// TIA Portal V19 export
FUNCTION "MB_VFD" : Void   // FC1, LAD
{ S7_Optimized_Access := 'TRUE' }
// stored: SetENOAutomatically false
   VAR_TEMP   // added for the SCL form of the ladder/FBD networks
      _w1 : Bool;
   END_VAR
BEGIN

REGION Network 1
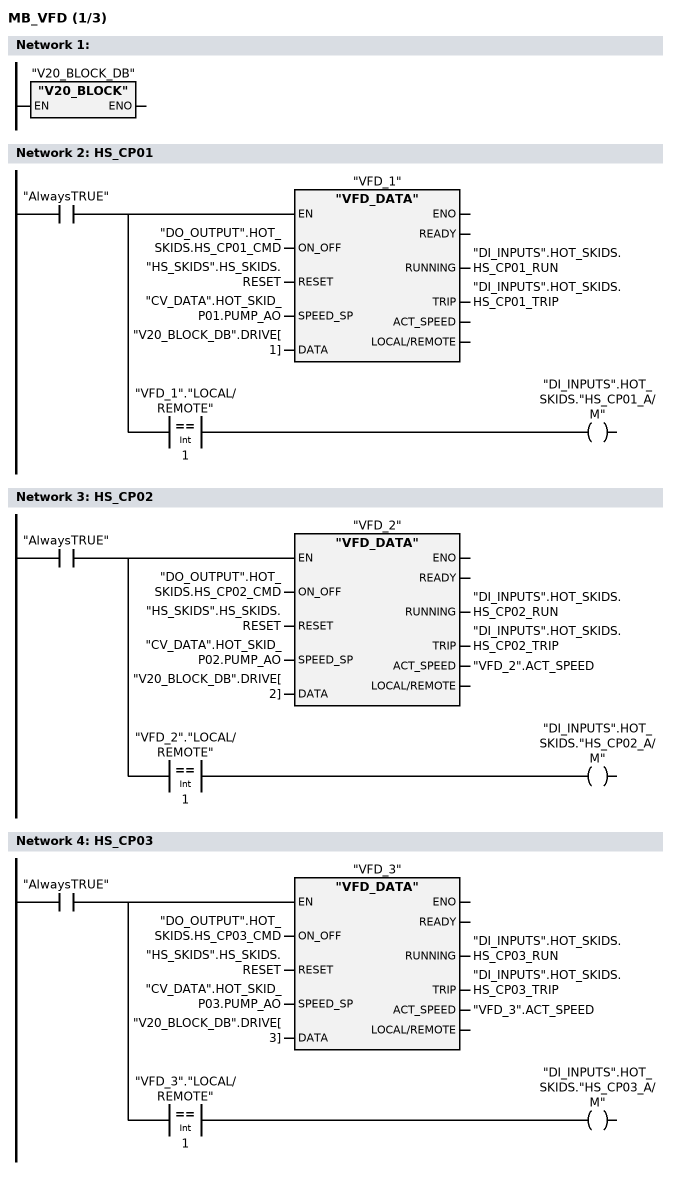
   RUNG wire#powerrail
      "V20_BLOCK_DB"()
   END_RUNG
   // the same network as SCL:
   "V20_BLOCK_DB"();   // "V20_BLOCK"
END_REGION

REGION Network 2: HS_CP01
   RUNG wire#powerrail
      Contact( "AlwaysTRUE" )
      wire#w1
      "VFD_1"(ON_OFF := "DO_OUTPUT".HOT_SKIDS.HS_CP01_CMD, RESET := "HS_SKIDS".HS_SKIDS.RESET, SPEED_SP := "CV_DATA".HOT_SKID_P01.PUMP_AO, DATA := "V20_BLOCK_DB".DRIVE[1], READY =>, RUNNING => "DI_INPUTS".HOT_SKIDS.HS_CP01_RUN, TRIP => "DI_INPUTS".HOT_SKIDS.HS_CP01_TRIP, ACT_SPEED =>, "LOCAL/REMOTE" =>)
   END_RUNG
   RUNG wire#w1
      { S7_Templates := "SrcType := Int" } EQ_Contact(in1 := "VFD_1"."LOCAL/REMOTE", in2 := 1)
      Coil( "DI_INPUTS".HOT_SKIDS."HS_CP01_A/M" )
   END_RUNG
   // the same network as SCL:
   #_w1 := "AlwaysTRUE";
   IF #_w1 THEN
       "VFD_1"(ON_OFF := "DO_OUTPUT".HOT_SKIDS.HS_CP01_CMD,   // "VFD_DATA"
               RESET := "HS_SKIDS".HS_SKIDS.RESET,
               SPEED_SP := "CV_DATA".HOT_SKID_P01.PUMP_AO,
               DATA := "V20_BLOCK_DB".DRIVE[1],
               RUNNING => "DI_INPUTS".HOT_SKIDS.HS_CP01_RUN,
               TRIP => "DI_INPUTS".HOT_SKIDS.HS_CP01_TRIP);
   END_IF;
   "DI_INPUTS".HOT_SKIDS."HS_CP01_A/M" := #_w1 AND ("VFD_1"."LOCAL/REMOTE" = 1);
END_REGION

REGION Network 3: HS_CP02
   RUNG wire#powerrail
      Contact( "AlwaysTRUE" )
      wire#w1
      "VFD_2"(ON_OFF := "DO_OUTPUT".HOT_SKIDS.HS_CP02_CMD, RESET := "HS_SKIDS".HS_SKIDS.RESET, SPEED_SP := "CV_DATA".HOT_SKID_P02.PUMP_AO, DATA := "V20_BLOCK_DB".DRIVE[2], READY =>, RUNNING => "DI_INPUTS".HOT_SKIDS.HS_CP02_RUN, TRIP => "DI_INPUTS".HOT_SKIDS.HS_CP02_TRIP, ACT_SPEED => "VFD_2".ACT_SPEED, "LOCAL/REMOTE" =>)
   END_RUNG
   RUNG wire#w1
      { S7_Templates := "SrcType := Int" } EQ_Contact(in1 := "VFD_2"."LOCAL/REMOTE", in2 := 1)
      Coil( "DI_INPUTS".HOT_SKIDS."HS_CP02_A/M" )
   END_RUNG
   // the same network as SCL:
   #_w1 := "AlwaysTRUE";
   IF #_w1 THEN
       "VFD_2"(ON_OFF := "DO_OUTPUT".HOT_SKIDS.HS_CP02_CMD,   // "VFD_DATA"
               RESET := "HS_SKIDS".HS_SKIDS.RESET,
               SPEED_SP := "CV_DATA".HOT_SKID_P02.PUMP_AO,
               DATA := "V20_BLOCK_DB".DRIVE[2],
               RUNNING => "DI_INPUTS".HOT_SKIDS.HS_CP02_RUN,
               TRIP => "DI_INPUTS".HOT_SKIDS.HS_CP02_TRIP,
               ACT_SPEED => "VFD_2".ACT_SPEED);
   END_IF;
   "DI_INPUTS".HOT_SKIDS."HS_CP02_A/M" := #_w1 AND ("VFD_2"."LOCAL/REMOTE" = 1);
END_REGION

REGION Network 4: HS_CP03
   RUNG wire#powerrail
      Contact( "AlwaysTRUE" )
      wire#w1
      "VFD_3"(ON_OFF := "DO_OUTPUT".HOT_SKIDS.HS_CP03_CMD, RESET := "HS_SKIDS".HS_SKIDS.RESET, SPEED_SP := "CV_DATA".HOT_SKID_P03.PUMP_AO, DATA := "V20_BLOCK_DB".DRIVE[3], READY =>, RUNNING => "DI_INPUTS".HOT_SKIDS.HS_CP03_RUN, TRIP => "DI_INPUTS".HOT_SKIDS.HS_CP03_TRIP, ACT_SPEED => "VFD_3".ACT_SPEED, "LOCAL/REMOTE" =>)
   END_RUNG
   RUNG wire#w1
      { S7_Templates := "SrcType := Int" } EQ_Contact(in1 := "VFD_3"."LOCAL/REMOTE", in2 := 1)
      Coil( "DI_INPUTS".HOT_SKIDS."HS_CP03_A/M" )
   END_RUNG
   // the same network as SCL:
   #_w1 := "AlwaysTRUE";
   IF #_w1 THEN
       "VFD_3"(ON_OFF := "DO_OUTPUT".HOT_SKIDS.HS_CP03_CMD,   // "VFD_DATA"
               RESET := "HS_SKIDS".HS_SKIDS.RESET,
               SPEED_SP := "CV_DATA".HOT_SKID_P03.PUMP_AO,
               DATA := "V20_BLOCK_DB".DRIVE[3],
               RUNNING => "DI_INPUTS".HOT_SKIDS.HS_CP03_RUN,
               TRIP => "DI_INPUTS".HOT_SKIDS.HS_CP03_TRIP,
               ACT_SPEED => "VFD_3".ACT_SPEED);
   END_IF;
   "DI_INPUTS".HOT_SKIDS."HS_CP03_A/M" := #_w1 AND ("VFD_3"."LOCAL/REMOTE" = 1);
END_REGION

REGION Network 5: CHS_CP01
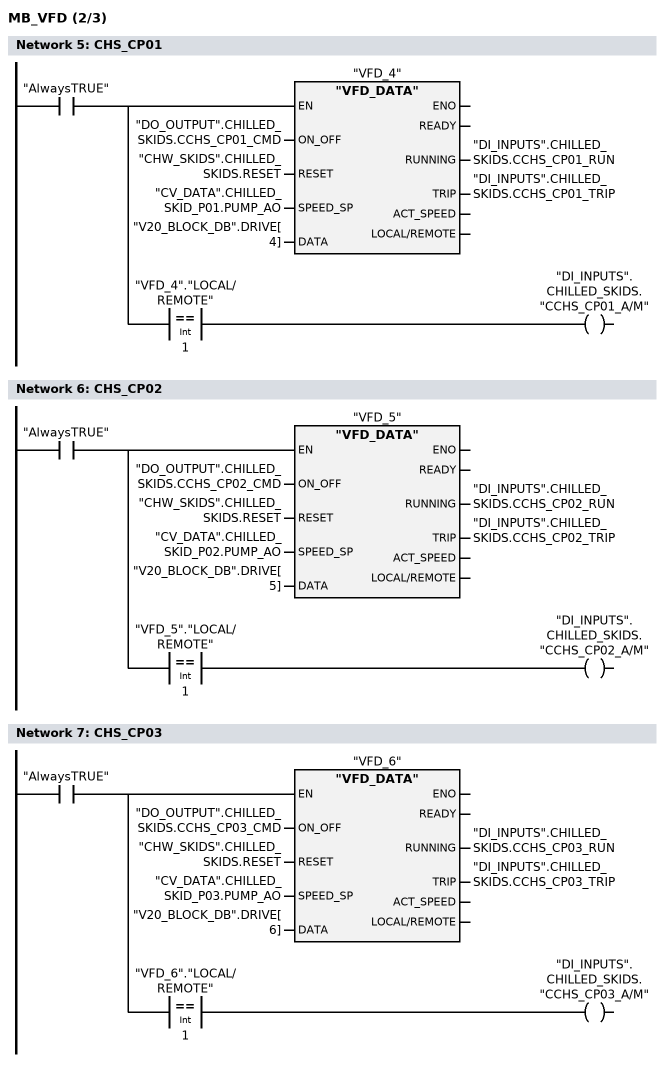
   RUNG wire#powerrail
      Contact( "AlwaysTRUE" )
      wire#w1
      "VFD_4"(ON_OFF := "DO_OUTPUT".CHILLED_SKIDS.CCHS_CP01_CMD, RESET := "CHW_SKIDS".CHILLED_SKIDS.RESET, SPEED_SP := "CV_DATA".CHILLED_SKID_P01.PUMP_AO, DATA := "V20_BLOCK_DB".DRIVE[4], READY =>, RUNNING => "DI_INPUTS".CHILLED_SKIDS.CCHS_CP01_RUN, TRIP => "DI_INPUTS".CHILLED_SKIDS.CCHS_CP01_TRIP, ACT_SPEED =>, "LOCAL/REMOTE" =>)
   END_RUNG
   RUNG wire#w1
      { S7_Templates := "SrcType := Int" } EQ_Contact(in1 := "VFD_4"."LOCAL/REMOTE", in2 := 1)
      Coil( "DI_INPUTS".CHILLED_SKIDS."CCHS_CP01_A/M" )
   END_RUNG
   // the same network as SCL:
   #_w1 := "AlwaysTRUE";
   IF #_w1 THEN
       "VFD_4"(ON_OFF := "DO_OUTPUT".CHILLED_SKIDS.CCHS_CP01_CMD,   // "VFD_DATA"
               RESET := "CHW_SKIDS".CHILLED_SKIDS.RESET,
               SPEED_SP := "CV_DATA".CHILLED_SKID_P01.PUMP_AO,
               DATA := "V20_BLOCK_DB".DRIVE[4],
               RUNNING => "DI_INPUTS".CHILLED_SKIDS.CCHS_CP01_RUN,
               TRIP => "DI_INPUTS".CHILLED_SKIDS.CCHS_CP01_TRIP);
   END_IF;
   "DI_INPUTS".CHILLED_SKIDS."CCHS_CP01_A/M" := #_w1 AND ("VFD_4"."LOCAL/REMOTE" = 1);
END_REGION

REGION Network 6: CHS_CP02
   RUNG wire#powerrail
      Contact( "AlwaysTRUE" )
      wire#w1
      "VFD_5"(ON_OFF := "DO_OUTPUT".CHILLED_SKIDS.CCHS_CP02_CMD, RESET := "CHW_SKIDS".CHILLED_SKIDS.RESET, SPEED_SP := "CV_DATA".CHILLED_SKID_P02.PUMP_AO, DATA := "V20_BLOCK_DB".DRIVE[5], READY =>, RUNNING => "DI_INPUTS".CHILLED_SKIDS.CCHS_CP02_RUN, TRIP => "DI_INPUTS".CHILLED_SKIDS.CCHS_CP02_TRIP, ACT_SPEED =>, "LOCAL/REMOTE" =>)
   END_RUNG
   RUNG wire#w1
      { S7_Templates := "SrcType := Int" } EQ_Contact(in1 := "VFD_5"."LOCAL/REMOTE", in2 := 1)
      Coil( "DI_INPUTS".CHILLED_SKIDS."CCHS_CP02_A/M" )
   END_RUNG
   // the same network as SCL:
   #_w1 := "AlwaysTRUE";
   IF #_w1 THEN
       "VFD_5"(ON_OFF := "DO_OUTPUT".CHILLED_SKIDS.CCHS_CP02_CMD,   // "VFD_DATA"
               RESET := "CHW_SKIDS".CHILLED_SKIDS.RESET,
               SPEED_SP := "CV_DATA".CHILLED_SKID_P02.PUMP_AO,
               DATA := "V20_BLOCK_DB".DRIVE[5],
               RUNNING => "DI_INPUTS".CHILLED_SKIDS.CCHS_CP02_RUN,
               TRIP => "DI_INPUTS".CHILLED_SKIDS.CCHS_CP02_TRIP);
   END_IF;
   "DI_INPUTS".CHILLED_SKIDS."CCHS_CP02_A/M" := #_w1 AND ("VFD_5"."LOCAL/REMOTE" = 1);
END_REGION

REGION Network 7: CHS_CP03
   RUNG wire#powerrail
      Contact( "AlwaysTRUE" )
      wire#w1
      "VFD_6"(ON_OFF := "DO_OUTPUT".CHILLED_SKIDS.CCHS_CP03_CMD, RESET := "CHW_SKIDS".CHILLED_SKIDS.RESET, SPEED_SP := "CV_DATA".CHILLED_SKID_P03.PUMP_AO, DATA := "V20_BLOCK_DB".DRIVE[6], READY =>, RUNNING => "DI_INPUTS".CHILLED_SKIDS.CCHS_CP03_RUN, TRIP => "DI_INPUTS".CHILLED_SKIDS.CCHS_CP03_TRIP, ACT_SPEED =>, "LOCAL/REMOTE" =>)
   END_RUNG
   RUNG wire#w1
      { S7_Templates := "SrcType := Int" } EQ_Contact(in1 := "VFD_6"."LOCAL/REMOTE", in2 := 1)
      Coil( "DI_INPUTS".CHILLED_SKIDS."CCHS_CP03_A/M" )
   END_RUNG
   // the same network as SCL:
   #_w1 := "AlwaysTRUE";
   IF #_w1 THEN
       "VFD_6"(ON_OFF := "DO_OUTPUT".CHILLED_SKIDS.CCHS_CP03_CMD,   // "VFD_DATA"
               RESET := "CHW_SKIDS".CHILLED_SKIDS.RESET,
               SPEED_SP := "CV_DATA".CHILLED_SKID_P03.PUMP_AO,
               DATA := "V20_BLOCK_DB".DRIVE[6],
               RUNNING => "DI_INPUTS".CHILLED_SKIDS.CCHS_CP03_RUN,
               TRIP => "DI_INPUTS".CHILLED_SKIDS.CCHS_CP03_TRIP);
   END_IF;
   "DI_INPUTS".CHILLED_SKIDS."CCHS_CP03_A/M" := #_w1 AND ("VFD_6"."LOCAL/REMOTE" = 1);
END_REGION

REGION Network 8: UCHS_CP01
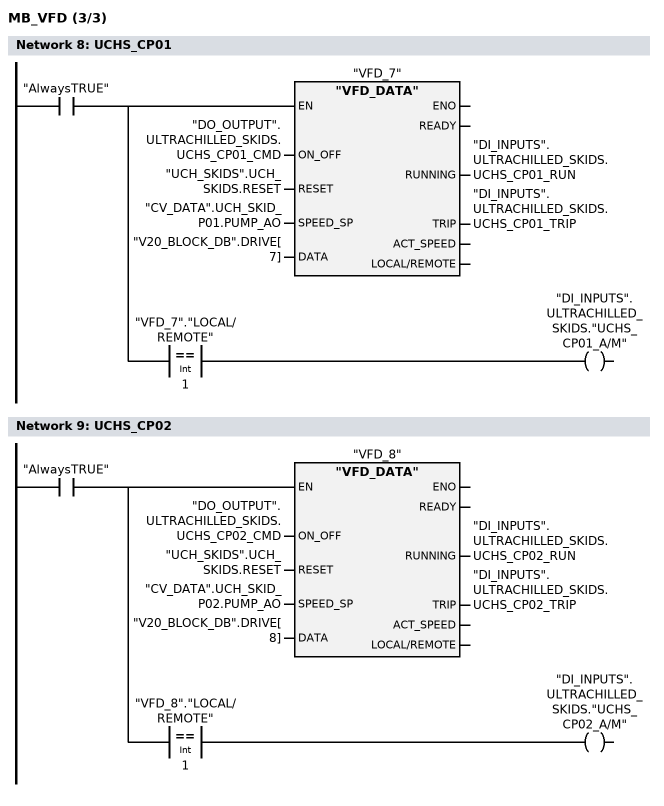
   RUNG wire#powerrail
      Contact( "AlwaysTRUE" )
      wire#w1
      "VFD_7"(ON_OFF := "DO_OUTPUT".ULTRACHILLED_SKIDS.UCHS_CP01_CMD, RESET := "UCH_SKIDS".UCH_SKIDS.RESET, SPEED_SP := "CV_DATA".UCH_SKID_P01.PUMP_AO, DATA := "V20_BLOCK_DB".DRIVE[7], READY =>, RUNNING => "DI_INPUTS".ULTRACHILLED_SKIDS.UCHS_CP01_RUN, TRIP => "DI_INPUTS".ULTRACHILLED_SKIDS.UCHS_CP01_TRIP, ACT_SPEED =>, "LOCAL/REMOTE" =>)
   END_RUNG
   RUNG wire#w1
      { S7_Templates := "SrcType := Int" } EQ_Contact(in1 := "VFD_7"."LOCAL/REMOTE", in2 := 1)
      Coil( "DI_INPUTS".ULTRACHILLED_SKIDS."UCHS_CP01_A/M" )
   END_RUNG
   // the same network as SCL:
   #_w1 := "AlwaysTRUE";
   IF #_w1 THEN
       "VFD_7"(ON_OFF := "DO_OUTPUT".ULTRACHILLED_SKIDS.UCHS_CP01_CMD,   // "VFD_DATA"
               RESET := "UCH_SKIDS".UCH_SKIDS.RESET,
               SPEED_SP := "CV_DATA".UCH_SKID_P01.PUMP_AO,
               DATA := "V20_BLOCK_DB".DRIVE[7],
               RUNNING => "DI_INPUTS".ULTRACHILLED_SKIDS.UCHS_CP01_RUN,
               TRIP => "DI_INPUTS".ULTRACHILLED_SKIDS.UCHS_CP01_TRIP);
   END_IF;
   "DI_INPUTS".ULTRACHILLED_SKIDS."UCHS_CP01_A/M" := #_w1 AND ("VFD_7"."LOCAL/REMOTE" = 1);
END_REGION

REGION Network 9: UCHS_CP02
   RUNG wire#powerrail
      Contact( "AlwaysTRUE" )
      wire#w1
      "VFD_8"(ON_OFF := "DO_OUTPUT".ULTRACHILLED_SKIDS.UCHS_CP02_CMD, RESET := "UCH_SKIDS".UCH_SKIDS.RESET, SPEED_SP := "CV_DATA".UCH_SKID_P02.PUMP_AO, DATA := "V20_BLOCK_DB".DRIVE[8], READY =>, RUNNING => "DI_INPUTS".ULTRACHILLED_SKIDS.UCHS_CP02_RUN, TRIP => "DI_INPUTS".ULTRACHILLED_SKIDS.UCHS_CP02_TRIP, ACT_SPEED =>, "LOCAL/REMOTE" =>)
   END_RUNG
   RUNG wire#w1
      { S7_Templates := "SrcType := Int" } EQ_Contact(in1 := "VFD_8"."LOCAL/REMOTE", in2 := 1)
      Coil( "DI_INPUTS".ULTRACHILLED_SKIDS."UCHS_CP02_A/M" )
   END_RUNG
   // the same network as SCL:
   #_w1 := "AlwaysTRUE";
   IF #_w1 THEN
       "VFD_8"(ON_OFF := "DO_OUTPUT".ULTRACHILLED_SKIDS.UCHS_CP02_CMD,   // "VFD_DATA"
               RESET := "UCH_SKIDS".UCH_SKIDS.RESET,
               SPEED_SP := "CV_DATA".UCH_SKID_P02.PUMP_AO,
               DATA := "V20_BLOCK_DB".DRIVE[8],
               RUNNING => "DI_INPUTS".ULTRACHILLED_SKIDS.UCHS_CP02_RUN,
               TRIP => "DI_INPUTS".ULTRACHILLED_SKIDS.UCHS_CP02_TRIP);
   END_IF;
   "DI_INPUTS".ULTRACHILLED_SKIDS."UCHS_CP02_A/M" := #_w1 AND ("VFD_8"."LOCAL/REMOTE" = 1);
END_REGION
END_FUNCTION
